FUNCTION_BLOCK FB_Machine EXTENDS FB_Module
(*
	Top-level module. Starting/stopping the machine starts/stops both stations.
	Start/stop/reset from the HMI with ocmd, or over MQTT (see cfgMqtt.enableRemoteCommands).
*)
VAR_INPUT
	(* Stations
	----------------------------------------------------------------------------------------------------*)
	{attribute 'OPC.UA.DA' := '1'}
	exampleStation		: FB_ExampleStation;
	{attribute 'OPC.UA.DA' := '1'}
	dosingStation		: FB_DosingStation; //ratio control loop example
	
	(* Communication
	----------------------------------------------------------------------------------------------------*)
	{attribute 'OPC.UA.DA' := '1'}
	{attribute 'OPC.UA.DA.StructuredType' := '1'}
	cfgMqtt				: ST_MqttConfiguration; //MQTT configuration
END_VAR
VAR
	{attribute 'OPC.UA.DA' := '0'} // internal MQTT client holds pointers OPC UA can't publish; status is in cfgMqtt/dashboard
	mqtt				: FB_MqttStatePublisher; //MQTT state publisher
END_VAR

SUPER^();

Stations();
Permissives();
Communication();

METHOD PROTECTED Communication
mqtt(cfg 			:= cfgMqtt,
	 machineState 	:= sts.State,
	 cycleCount 	:= exampleStation.stsStation.cycleCount);

//Remote commands are handled like program commands
IF mqtt.cmd <> E_ModuleCommand.None THEN
	pcmd := mqtt.cmd;
END_IF
END_METHOD

METHOD PROTECTED Permissives //set module permissives and interlocks
//Started once every station is running
PermStartComplete.cfg.condText[0] := 'Example station started';
PermStartComplete.cfg.condText[1] := 'Dosing station started';
PermStartComplete.perm.0 := exampleStation.sts.Started;
PermStartComplete.perm.1 := dosingStation.sts.Started;

//Stopped once every station is stopped
PermStopComplete.cfg.condText[0] := 'Example station stopped';
PermStopComplete.cfg.condText[1] := 'Dosing station stopped';
PermStopComplete.perm.0 := exampleStation.sts.Stopped;
PermStopComplete.perm.1 := dosingStation.sts.Stopped;

//A faulted station stops the machine
IntlkAuto.cfg.condText[0] := 'Example station not faulted';
IntlkAuto.cfg.condText[1] := 'Dosing station not faulted';
IntlkAuto.perm.0 := NOT exampleStation.sts.Faulted;
IntlkAuto.perm.1 := NOT dosingStation.sts.Faulted;
END_METHOD

METHOD PUBLIC Reset : BOOL
exampleStation.cmdReset := TRUE;
dosingStation.cmdReset := TRUE;
Reset := TRUE;
END_METHOD

METHOD PROTECTED Started : BOOL
//Stations run their own sequences while the machine is started
END_METHOD

METHOD PROTECTED Starting : BOOL
exampleStation.pcmd := E_ModuleCommand.Start;
dosingStation.pcmd := E_ModuleCommand.Start;
END_METHOD

METHOD PROTECTED Stations //call child modules
exampleStation();
dosingStation();

inpChildFaulted := exampleStation.sts.Faulted OR dosingStation.sts.Faulted;
END_METHOD

METHOD PROTECTED Stopping : BOOL
exampleStation.pcmd := E_ModuleCommand.Stop;
dosingStation.pcmd := E_ModuleCommand.Stop;
END_METHOD

END_FUNCTION_BLOCK

(* stored: Version 1.1.0.1, ProductVersion 3.1.4024.12
   POU FB_Machine: Id {fd543e1c-2eca-4831-ae5c-5f1ac010e45e}, SpecialFunc None
   Folder Protected: Id {58843e9d-4289-4344-8d11-03266e1b722a}
   Folder Logic: Id {3f3dc444-fa34-4e97-be9c-d57c389576f9}
   Folder States: Id {b6dfe07d-6d5d-45af-b0bd-12d2473dfa3a}
   Folder Public: Id {a4c667e2-6e19-4bc0-b242-943d38308146}
   Folder Control: Id {5ed18d35-54a8-436a-91d5-f96cb2f8da01}
   Method Communication: Id {e2b37e0b-5eb1-4160-9702-ac335e75a9a8}
   Method Permissives: Id {1d31ecc1-e23a-4b40-80b2-f8cf2e2bed17}
   Method Reset: Id {cb192e32-b467-40eb-bce0-ecf1ba70a10f}
   Method Started: Id {6572cca9-89d7-4580-ba96-befb8e702fef}
   Method Starting: Id {a1a124df-8592-4282-a52c-e0737dc46e9e}
   Method Stations: Id {28a083f7-7251-46a3-abba-099a8be6f6ae}
   Method Stopping: Id {daf1d2a3-6b3e-4e18-a0d6-7c6c58ffd8ee} *)
